(* IEC 61131-3 sources: plcassist-cli/packages/volt-lsp-iec/test-corpus/pro2193/Device/Plc Logic/Application/09 Misc/Library Manager/CAA SegBufMan, 37 files *)

(* ---- RSHANDLING.gvl ---- *)
VAR_GLOBAL
	G_BUFFERCLASS : BufferClass;
	G_QUEUECLASS : QueueClass;
END_VAR

(* ---- VERSIONCONSTANTS.gvl ---- *)
VAR_GLOBAL
	GC_BYVERSION : BYTE := 1;
	GC_BYVERSION_1 : BYTE := 0;
END_VAR

(* ---- _BUFFERADDREF.fun ---- *)
FUNCTION _BUFFERADDREF : ERROR
VAR_INPUT
	HBUFFER : CAA.HANDLE;
END_VAR
END_FUNCTION

(* ---- _CHAINBUFFER.fun ---- *)
FUNCTION _CHAINBUFFER : CAA.HANDLE
VAR_INPUT
	HHEAD : CAA.HANDLE;
	HTAIL : CAA.HANDLE;
	PEERROR : POINTER TO ERROR;
END_VAR
END_FUNCTION

(* ---- _COPYBUFFERDATA.fun ---- *)
FUNCTION _COPYBUFFERDATA : ERROR
VAR_INPUT
	HBUFFER : CAA.HANDLE;
	SZOFFSET : CAA.SIZE;
	SZLENGTH : CAA.SIZE;
	PDATA : CAA.PVOID;
	SZSIZE : CAA.SIZE;
END_VAR
END_FUNCTION

(* ---- _CREATEBUFFER.fun ---- *)
FUNCTION _CREATEBUFFER : CAA.HANDLE
VAR_INPUT
	SZSIZE : CAA.SIZE;
	PDATA : CAA.PVOID;
	XPERMANENT : BOOL;
	PEERROR : POINTER TO ERROR;
END_VAR
END_FUNCTION

(* ---- _CREATEQUEUE.fun ---- *)
FUNCTION _CREATEQUEUE : CAA.HANDLE
VAR_INPUT
	PEERROR : POINTER TO ERROR;
END_VAR
END_FUNCTION

(* ---- _DELETEBUFFER.fun ---- *)
FUNCTION _DELETEBUFFER : ERROR
VAR_INPUT
	HBUFFER : CAA.HANDLE;
END_VAR
END_FUNCTION

(* ---- _DELETEQUEUE.fun ---- *)
FUNCTION _DELETEQUEUE : ERROR
VAR_INPUT
	HQUEUE : CAA.HANDLE;
END_VAR
END_FUNCTION

(* ---- _DEQUEUEBUFFER.fun ---- *)
FUNCTION _DEQUEUEBUFFER : CAA.HANDLE
VAR_INPUT
	HQUEUE : CAA.HANDLE;
	PEERROR : POINTER TO ERROR;
END_VAR
END_FUNCTION

(* ---- _ENQUEUEBUFFER.fun ---- *)
FUNCTION _ENQUEUEBUFFER : ERROR
VAR_INPUT
	HQUEUE : CAA.HANDLE;
	HBUFFER : CAA.HANDLE;
END_VAR
END_FUNCTION

(* ---- _GETBUFFERSIZE.fun ---- *)
FUNCTION _GETBUFFERSIZE : CAA.SIZE
VAR_INPUT
	HBUFFER : CAA.HANDLE;
	PEERROR : POINTER TO ERROR;
END_VAR
END_FUNCTION

(* ---- _GETQUEUELENGTH.fun ---- *)
FUNCTION _GETQUEUELENGTH : CAA.SIZE
VAR_INPUT
	HQUEUE : CAA.HANDLE;
	PEERROR : POINTER TO ERROR;
END_VAR
END_FUNCTION

(* ---- _GETSEGMENTDATAPOINTER.fun ---- *)
FUNCTION _GETSEGMENTDATAPOINTER : CAA.PVOID
VAR_INPUT
	HBUFFER : CAA.HANDLE;
	PSZSIZE : POINTER TO CAA.SIZE;
	PXPERMANENT : POINTER TO BOOL;
	PEERROR : POINTER TO ERROR;
END_VAR
END_FUNCTION

(* ---- _MOVETOBUFFEROFFSET.fun ---- *)
FUNCTION _MOVETOBUFFEROFFSET : ERROR
VAR_INPUT
	HBUFFER : CAA.HANDLE;
	SZOFFSET : CAA.SIZE;
END_VAR
END_FUNCTION

(* ---- _MOVETONEXTSEGMENT.fun ---- *)
FUNCTION _MOVETONEXTSEGMENT : ERROR
VAR_INPUT
	HBUFFER : CAA.HANDLE;
END_VAR
END_FUNCTION

(* ---- _SLICEBUFFER.fun ---- *)
FUNCTION _SLICEBUFFER : CAA.HANDLE
VAR_INPUT
	HBUFFER : CAA.HANDLE;
	SZOFFSET : CAA.SIZE;
	SZLENGTH : CAA.SIZE;
	PEERROR : POINTER TO ERROR;
END_VAR
END_FUNCTION

(* ---- CHAINBUFFER.fun ---- *)
FUNCTION CHAINBUFFER : CAA.HANDLE
VAR_INPUT
	HHEAD : CAA.HANDLE;
	HTAIL : CAA.HANDLE;
	PEERROR : POINTER TO ERROR;
END_VAR
END_FUNCTION

(* ---- COPYBUFFERDATA.fun ---- *)
FUNCTION COPYBUFFERDATA : ERROR
VAR_INPUT
	HBUFFER : CAA.HANDLE;
	SZOFFSET : CAA.SIZE;
	SZLENGTH : CAA.SIZE;
	PDATA : CAA.PVOID;
	SZSIZE : CAA.SIZE;
END_VAR
END_FUNCTION

(* ---- CREATEBUFFER.fun ---- *)
FUNCTION CREATEBUFFER : CAA.HANDLE
VAR_INPUT
	SZSIZE : CAA.SIZE;
	PDATA : CAA.PVOID;
	XPERMANENT : BOOL;
	PEERROR : POINTER TO ERROR;
END_VAR
END_FUNCTION

(* ---- CREATEQUEUE.fun ---- *)
FUNCTION CREATEQUEUE : CAA.HANDLE
VAR_INPUT
	PEERROR : POINTER TO ERROR;
END_VAR
END_FUNCTION

(* ---- DELETEBUFFER.fun ---- *)
FUNCTION DELETEBUFFER : ERROR
VAR_INPUT
	HBUFFER : CAA.HANDLE;
END_VAR
END_FUNCTION

(* ---- DELETEQUEUE.fun ---- *)
FUNCTION DELETEQUEUE : ERROR
VAR_INPUT
	HQUEUE : CAA.HANDLE;
END_VAR
END_FUNCTION

(* ---- DEQUEUEBUFFER.fun ---- *)
FUNCTION DEQUEUEBUFFER : CAA.HANDLE
VAR_INPUT
	HQUEUE : CAA.HANDLE;
	PEERROR : POINTER TO ERROR;
END_VAR
END_FUNCTION

(* ---- ENQUEUEBUFFER.fun ---- *)
FUNCTION ENQUEUEBUFFER : ERROR
VAR_INPUT
	HQUEUE : CAA.HANDLE;
	HBUFFER : CAA.HANDLE;
END_VAR
END_FUNCTION

(* ---- GETBUFFERSIZE.fun ---- *)
FUNCTION GETBUFFERSIZE : CAA.SIZE
VAR_INPUT
	HBUFFER : CAA.HANDLE;
	PEERROR : POINTER TO ERROR;
END_VAR
END_FUNCTION

(* ---- GETLIBVERSION.fun ---- *)
FUNCTION GETLIBVERSION : VERSION
END_FUNCTION

(* ---- GETLIBVERSIONNUMBER.fun ---- *)
FUNCTION GETLIBVERSIONNUMBER : DWORD
END_FUNCTION

(* ---- GETQUEUELENGTH.fun ---- *)
FUNCTION GETQUEUELENGTH : CAA.SIZE
VAR_INPUT
	HQUEUE : CAA.HANDLE;
	PEERROR : POINTER TO ERROR;
END_VAR
END_FUNCTION

(* ---- GETSEGMENTDATAPOINTER.fun ---- *)
FUNCTION GETSEGMENTDATAPOINTER : CAA.PVOID
VAR_INPUT
	HBUFFER : CAA.HANDLE;
	PSZSIZE : POINTER TO CAA.SIZE;
	PXPERMANENT : POINTER TO BOOL;
	PEERROR : POINTER TO ERROR;
END_VAR
END_FUNCTION

(* ---- GETSUPPLIERVERSION.fun ---- *)
FUNCTION GETSUPPLIERVERSION : WORD
VAR_INPUT
	XDUMMY : BOOL;
END_VAR
END_FUNCTION

(* ---- ISLIBRELEASED.fun ---- *)
FUNCTION ISLIBRELEASED : BOOL
END_FUNCTION

(* ---- MOVETOBUFFEROFFSET.fun ---- *)
FUNCTION MOVETOBUFFEROFFSET : ERROR
VAR_INPUT
	HBUFFER : CAA.HANDLE;
	SZOFFSET : CAA.SIZE;
END_VAR
END_FUNCTION

(* ---- MOVETONEXTSEGMENT.fun ---- *)
FUNCTION MOVETONEXTSEGMENT : ERROR
VAR_INPUT
	HBUFFER : CAA.HANDLE;
END_VAR
END_FUNCTION

(* ---- SLICEBUFFER.fun ---- *)
FUNCTION SLICEBUFFER : CAA.HANDLE
VAR_INPUT
	HBUFFER : CAA.HANDLE;
	SZOFFSET : CAA.SIZE;
	SZLENGTH : CAA.SIZE;
	PEERROR : POINTER TO ERROR;
END_VAR
END_FUNCTION

(* ---- BUFFERCLASS.fb ---- *)
FUNCTION_BLOCK BUFFERCLASS EXTENDS RSMClass
END_FUNCTION_BLOCK

METHOD CLOSE : RSM.ERROR
VAR_INPUT
	HHANDLE : CAA.HANDLE;
END_VAR
END_METHOD

(* ---- QUEUECLASS.fb ---- *)
FUNCTION_BLOCK QUEUECLASS EXTENDS RSMClass
END_FUNCTION_BLOCK

METHOD CLOSE : RSM.ERROR
VAR_INPUT
	HHANDLE : CAA.HANDLE;
END_VAR
END_METHOD
